(* IEC 61131-3 sources: trust-platform/examples/hardware_8do/src, 2 files *)

(* ---- config.st ---- *)
CONFIGURATION Config
RESOURCE MainResource ON PLC
    TASK MainTask (INTERVAL := T#10ms, PRIORITY := 1);
    PROGRAM P1 WITH MainTask : Main;
END_RESOURCE
VAR_CONFIG
    P1.DO0 AT %QX0.0 : BOOL;
    P1.DO1 AT %QX0.1 : BOOL;
    P1.DO2 AT %QX0.2 : BOOL;
    P1.DO3 AT %QX0.3 : BOOL;
    P1.DO4 AT %QX0.4 : BOOL;
    P1.DO5 AT %QX0.5 : BOOL;
    P1.DO6 AT %QX0.6 : BOOL;
    P1.DO7 AT %QX0.7 : BOOL;
END_VAR
END_CONFIGURATION

(* ---- Main.st ---- *)
(*
    Hardware Backend: 8 Digital Outputs

    This is a minimal ST program that defines I/O variables.

    The actual control logic can come from:
    - Blockly visual programs (interpreted via control endpoint)
    - Statechart programs (interpreted via control endpoint)
    - ST code written here

    For visual editors (Blockly/Statechart), the outputs are controlled
    through the control endpoint at /tmp/trust-debug.sock, not by this code.
*)

PROGRAM Main
VAR
    // Digital outputs mapped to hardware (EL2008 or GPIO)
    DO0 AT %QX0.0 : BOOL;
    DO1 AT %QX0.1 : BOOL;
    DO2 AT %QX0.2 : BOOL;
    DO3 AT %QX0.3 : BOOL;
    DO4 AT %QX0.4 : BOOL;
    DO5 AT %QX0.5 : BOOL;
    DO6 AT %QX0.6 : BOOL;
    DO7 AT %QX0.7 : BOOL;

    // Heartbeat to show program is running
    heartbeat : BOOL;
END_VAR

// Toggle heartbeat every cycle
heartbeat := NOT heartbeat;

// For visual editors: outputs controlled via control endpoint
// For ST programs: add your logic here

END_PROGRAM
